// TIA Portal V21 export
// export: Created 2026-11-08T19:42:57.5114689Z, ExportSetting WithDefaults, DisplayName Totally Integrated Automation Portal, DisplayVersion V21 Update 3, DisplayName STEP 7 Professional, DisplayVersion V21 Update 3, DisplayName STEP 7 Safety, DisplayVersion V21, DisplayName Tech WebApplication, DisplayVersion V21, DisplayName WinCC Basic/Comfort/Advanced, DisplayVersion V21 Update 3, DisplayName WinCC Unified, DisplayVersion V21 Update 3
VAR_GLOBAL   // PLC tag table "TagTable_1"
   Tag_Bool_1 AT %M0.0 : Bool;
   In_Bool AT %I0.1 : Bool;
   Out_Bool AT %Q2.0 : Bool;
   M_Int AT %MW20 : Int;
   M_Real AT %MD24 : Real;
   In_Word AT %IW4 : Word;
   Out_Byte AT %QB3 : Byte;
   M_DInt AT %MD28 : DInt;   // DInt Kommentar
   M_Time AT %MD32 : Time;
END_VAR
